(* IEC 61131-3 sources: Caravan/Archiv/12-04-19/Stations/MachineControl/MachineControl/Class/HmiTextList35, 1 file *)

(* ---- HmiTextList35.st ---- *)
(*!
<Class
	Name               = "HmiTextList35"
	Revision           = "0.1"
	RealtimeTask       = "false"
	CyclicTask         = "false"
	BackgroundTask     = "false"
	Sigmatek           = "true"
	OSInterface        = "false"
	HighPriority       = "false"
	Automatic          = "false"
	UpdateMode         = "Prescan"
	SharedCommandTable = "true"
	Objectsize         = "(284,120)">
	<Channels>
		<Server Name="ByteSize" Visualized="false" Initialize="false" WriteProtected="true" Retentive="false"/>
		<Server Name="ClassSvr" Visualized="false" Initialize="false" WriteProtected="true" Retentive="false"/>
	</Channels>
	<RevDoku>
		<Owner Company="sigmatek" Author="kolott"/>
		<Dokumentation Revision="0.1" Date="2014-03-28" Author="kolott" Company="sigmatek" Description="server ByteSize added"/>
	</RevDoku>
</Class>
*)
HmiTextList35 : CLASS
  //Servers:
	ClassSvr 	: SvrChCmd_UDINT;
	ByteSize 	: SvrCh_UDINT;
  //Clients:
  //Variables:
		Ptr 	: ^void;
		xData : ARRAY [0..20000] OF UINT;

		xOffset : ARRAY [0..5000] OF UDINT;

		xSize 	: UDINT;
  //Functions:

	FUNCTION GLOBAL End
		VAR_OUTPUT
			retcode 	: ^void;
		END_VAR;

	FUNCTION GLOBAL Free;

	FUNCTION GLOBAL Start;

	FUNCTION GLOBAL AddEntry
		VAR_INPUT
			txt 	: ^UINT;
		END_VAR
		VAR_OUTPUT
			retcode 	: UDINT;
		END_VAR;

	FUNCTION SeekText
		VAR_INPUT
			txt 	: ^UINT;
			length 	: UDINT;
		END_VAR
		VAR_OUTPUT
			retcode 	: UDINT;
		END_VAR;
  //Tables:
	FUNCTION @STD
		VAR_OUTPUT
			ret_code	: CONFSTATES;
		END_VAR;
	FUNCTION GLOBAL TAB @CT_;
END_CLASS;

#includeC "..\LseEasy\Create.h"

FUNCTION GLOBAL HmiTextList35::Free

  Start();

END_FUNCTION

FUNCTION GLOBAL HmiTextList35::Start

  xSize    := 0;
  Ptr      := NIL;
  ByteSize := 0;

END_FUNCTION

FUNCTION HmiTextList35::SeekText
  var_input
    txt : ^uint;
    length : udint;
  end_var
  var_output
    retcode : udint;
  end_var
  var
    ptl : ^_BOX_TEXTLIST;
    nox : udint;
    ph : ^uint;
  end_var

  ptl$^void := Ptr;

  if(ptl <> NIL) then
    nox := ptl^.no;
    while(nox) do
      nox -= 1;
      ph := #ptl^.data[0] + xOffset[nox];
      if(ph^ = txt^) then
        if(_memcmp(ph, txt, length) = 0) then
          retcode := nox;
          return;
        end_if;
      end_if;
    end_while;
  end_if;

  retcode := 16#FFFFFFFF;

END_FUNCTION

FUNCTION GLOBAL HmiTextList35::AddEntry
  var_input
    txt : ^uint;
  end_var
  var_output
    retcode : udint;
  end_var
  var
    ptl : ^_BOX_TEXTLIST;
    length : udint;
    ph : ^uint;
  end_var

  retcode := 16#FFFFFFFF;

  if(txt <> NIL) then
    if(Ptr = NIL) then
      xSize := 0;
      Ptr   := #xData[0];
      _memset(Ptr, 0, sizeof(xData));
      _memset(#xOffset[0], 16#FF, sizeof(xOffset));
      ptl$^void         := Ptr;
      ptl^.no           := 0;
      ptl^.boxhdr.size  := 0;
      ptl^.boxhdr.crc32 := 0;
    end_if;

    ptl$^void := Ptr;
    length    := StrLen3(txt) + 1;
    length    := length * 2;
    retcode   := SeekText(txt, length);

    if(retcode = 16#FFFFFFFF) then
      if((xSize + length) < (sizeof(xData) - sizeof(_BIGBOX_HEADER) - 4)) then
        ph               := #ptl^.data[0] + xSize;
        _memcpy(ph, txt, length);
        retcode          := ptl^.no;
        xOffset[retcode] := xSize;
        xSize            += length;
        ptl^.no          += 1;
      end_if;
    end_if;
  end_if;

END_FUNCTION

FUNCTION GLOBAL HmiTextList35::End
	VAR_OUTPUT
		retcode 	: ^void;
	END_VAR
  var
    ptl : ^_BOX_TEXTLIST;
  end_var

  if(Ptr <> NIL) then
    ptl$^void := Ptr;
    ClassSvr  := ptl^.no;
    ptl^.boxhdr.size := sizeof(ptl^.boxhdr) + sizeof(ptl^.no);
    end_BIGBOX_HEADER(#ptl^.boxhdr, xSize);
    ByteSize := ptl^.boxhdr.size;
  end_if;

  retcode := Ptr;

END_FUNCTION
